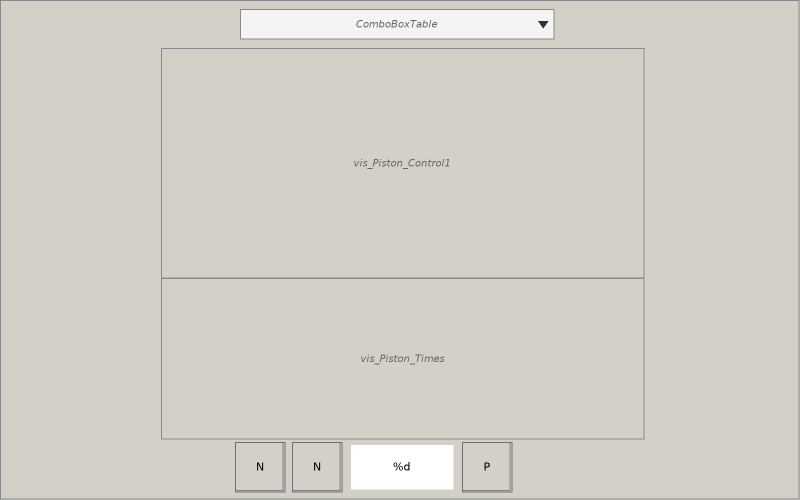
VISUALIZATION vis_Piston_Select_1  // 800x500
    Frame (161,48 483x230)
        shows vis_Piston_Control1(stPis := stPis[iPis_sel])
    Frame (161,278 483x161)
        shows vis_Piston_Times(stPis := stPis[iPis_sel])
    Button (292,442 50x50), "N"
        tap prg_Piston.bPis_Next_N
    Button (462,442 50x50), "P"
        tap prg_Piston.bPis_Next_P
    Textfield (350,444 104x46), "%d", text variable: iPis_sel
    ComboBoxTable (240,9 314x30), variable: iPis_sel, data array: arPisName
        p1128707560: C_MAX_Pistons_Exist
        p3854506369: arPisName[INDEX].Num
        p1892666644: arPisName[INDEX].Description
    Button (235,442 50x50), "N"
        tap prg_Piston.bPis_Next_N
END_VISUALIZATION

(* stored: Version 1.1.0.1, ProductVersion 3.1.4024.12
   Visu vis_Piston_Select_1: Id {ec812f09-9e9f-4579-84c4-a08a77964f1c} *)
